Fanuc KAREL source: KA00207.KL

PROGRAM KA00207
%NOLOCKGROUP
VAR
  SRC: ARRAY[4] OF VECTOR
  DST: ARRAY[4] OF JOINTPOS
BEGIN
  DST = SRC
END KA00207
